(* IEC 61131-3 sources: llm-plc-st-eval/data/processed_definitivo/qwen2.5-coder_14b/I4/zero_shot, 3 files *)

(* ---- ejec_1.st ---- *)
FUNCTION_BLOCK FB_EstrellaTriangulo
VAR_INPUT
    btnMarcha : BOOL; // Botón de marcha
    btnParo : BOOL;   // Botón de paro
END_VAR

VAR_OUTPUT
    kM : BOOL;       // Contactor principal
    kY : BOOL;       // Contactor de estrella
    kD : BOOL;       // Contactor de triángulo
END_VAR

VAR
    timerEstrella : TON; // Temporizador para el contacto de estrella
    timerMuerto : TON;   // Temporizador para el tiempo muerto
    estado : INT;       // Variable de estado del arranque
END_VAR

// Inicialización de temporizadores
timerEstrella(IN := FALSE, PT := T#8S);
timerMuerto(IN := FALSE, PT := T#100MS);

// Máquina de estados
CASE estado OF
    0: // Estado inicial
        IF btnMarcha THEN
            kM := TRUE; // Activar el contactor principal
            kY := TRUE; // Activar el contactor de estrella
            timerEstrella(IN := TRUE); // Iniciar temporizador para el contacto de estrella
            estado := 1; // Transición al estado 1
        END_IF

    1: // Esperando el fin del temporizador de estrella
        IF timerEstrella.Q THEN
            kY := FALSE; // Desactivar el contactor de estrella
            timerMuerto(IN := TRUE); // Iniciar temporizador para el tiempo muerto
            estado := 2; // Transición al estado 2
        END_IF

    2: // Esperando el fin del temporizador de tiempo muerto
        IF timerMuerto.Q THEN
            kD := TRUE; // Activar el contactor de triángulo
            estado := 3; // Transición al estado 3
        END_IF

    3: // Estado final
        // Mantener los contactores activados según el estado actual
        IF btnParo THEN
            kM := FALSE; // Desactivar el contactor principal
            kY := FALSE; // Desactivar el contactor de estrella
            kD := FALSE; // Desactivar el contactor de triángulo
            estado := 0; // Reiniciar a estado inicial
        END_IF
END_CASE

(* ---- ejec_2.st ---- *)
FUNCTION_BLOCK FB_EstrellaTriangulo
VAR_INPUT
    btnMarcha : BOOL; // Botón de marcha
    btnParo : BOOL; // Botón de paro
END_VAR

VAR_OUTPUT
    kM : BOOL; // Contactor principal
    kY : BOOL; // Contactor de estrella
    kD : BOOL; // Contactor de triángulo
END_VAR

VAR
    timerStar : TON; // Temporizador para el contacto de estrella
    timerDelta : TON; // Temporizador para el contacto de triángulo
    state : INT := 0; // Estado actual del programa
    deadTime : TON; // Temporizador para el tiempo muerto
END_VAR

// Inicialización de temporizadores
timerStar(IN := FALSE, PT := T#8S);
timerDelta(IN := FALSE, PT := T#100MS);
deadTime(IN := FALSE, PT := T#100MS);

// Lógica del programa
CASE state OF
    0: // Estado inicial
        IF btnMarcha THEN
            kM := TRUE;
            kY := TRUE;
            timerStar(IN := TRUE);
            state := 1;
        END_IF
        IF btnParo THEN
            kM := FALSE;
            kY := FALSE;
            kD := FALSE;
            state := 0;
        END_IF

    1: // Esperando para desactivar kY
        IF timerStar.Q THEN
            kY := FALSE;
            timerStar(IN := FALSE);
            deadTime(IN := TRUE);
            state := 2;
        END_IF
        IF btnParo THEN
            kM := FALSE;
            kY := FALSE;
            kD := FALSE;
            state := 0;
        END_IF

    2: // Tiempo muerto
        IF deadTime.Q THEN
            kD := TRUE;
            deadTime(IN := FALSE);
            state := 3;
        END_IF
        IF btnParo THEN
            kM := FALSE;
            kY := FALSE;
            kD := FALSE;
            state := 0;
        END_IF

    3: // Estado final
        IF btnParo THEN
            kM := FALSE;
            kY := FALSE;
            kD := FALSE;
            state := 0;
        END_IF
END_CASE

(* ---- ejec_3.st ---- *)
FUNCTION_BLOCK FB_EstrellaTriangulo
VAR_INPUT
    btnMarcha : BOOL; // Botón de marcha
    btnParo : BOOL;   // Botón de paro
END_VAR

VAR_OUTPUT
    kM : BOOL; // Contactor principal
    kY : BOOL; // Contactor de estrella
    kD : BOOL; // Contactor de triángulo
END_VAR

VAR
    timerEstrella : TON; // Temporizador para el contacto de estrella
    timerMuerto : TON;   // Temporizador para el tiempo muerto
    estado : INT;       // Estado actual del arranque estrella-triángulo
END_VAR

// Estados del arranque estrella-triángulo
CONST
    ESTADO_INICIAL := 0;
    ESTADO_MARCHA := 1;
    ESTADO_TIEMPO_MUERTO := 2;
    ESTADO_TRIANGULO := 3;
END_CONST

// Inicialización
IF NOT btnParo THEN
    CASE estado OF
        ESTADO_INICIAL:
            kM := FALSE;
            kY := FALSE;
            kD := FALSE;
            IF btnMarcha THEN
                estado := ESTADO_MARCHA;
                kM := TRUE;
                kY := TRUE;
                timerEstrella(IN := TRUE, PT := T#8S);
            END_IF;

        ESTADO_MARCHA:
            IF timerEstrella.Q THEN
                estado := ESTADO_TIEMPO_MUERTO;
                kY := FALSE;
                timerMuerto(IN := TRUE, PT := T#100MS);
            END_IF;

        ESTADO_TIEMPO_MUERTO:
            IF timerMuerto.Q THEN
                estado := ESTADO_TRIANGULO;
                kD := TRUE;
            END_IF;

        ESTADO_TRIANGULO:
            // Mantener kD activo mientras no se presione btnParo
            kD := TRUE;
    END_CASE;
ELSE
    // Paro forzado
    estado := ESTADO_INICIAL;
    kM := FALSE;
    kY := FALSE;
    kD := FALSE;
    timerEstrella(IN := FALSE);
    timerMuerto(IN := FALSE);
END_IF;
